(* IEC 61131-3 sources: Caravan/Archiv/12-04-19/Stations/Terminal/HMI/Network/IPCONF_IPConfigHMI, 1 file *)

(* ---- ONE_IPCONF_IPConfigHMI_Table.st ---- *)
#define OBJECTS_CONFIG

//Define part of class _IPConfigMain
//===========================================================================================================

#define MaxNoStations         50        // max. allowed No of stations

#define IPcfgWindowNrMsgBox   51000     // Window-Number of the Message Box

//===========================================================================================================
#include <.\LoaderItf.h>
//Define part of class _IPConfigStation
//===========================================================================================================

#define NiCmdIF_HmsWaitIF     20        // NewInst() command to IF object:
                                        // Time Delay for command work [100 ms] within the IF object

//===========================================================================================================

FUNCTION GLOBAL TAB ONE_IPCONF_IPConfigHMI
-1$UINT, 0$UINT,
0$UINT, 0$UINT,

13$UDINT,
TO_UDINT(3788417926), "_Global", 0$UINT, 14$UINT, 0$UINT,
TO_UDINT(1245802338), "_IPConfigIF", 1$UINT, 1$UINT, 1$UINT,
TO_UDINT(4058854491), "_IPConfigMain", 1$UINT, 2$UINT, 1$UINT,
TO_UDINT(148468755), "_IPConfigStation", 1$UINT, 2$UINT, 2$UINT,
TO_UDINT(4101473903), "_SearchUsbFiletoReset", 1$UINT, 0$UINT, 1$UINT,
TO_UDINT(2550379949), "Client_Splitter_10", 1$UINT, 2$UINT, 1$UINT,
TO_UDINT(1524808134), "Client_Splitter_Base", 1$UINT, 1$UINT, 0$UINT,
TO_UDINT(2225119864), "MerkerEx", 1$UINT, 21$UINT, 0$UINT,
TO_UDINT(3068426329), "NetworkConfig", 1$UINT, 31$UINT, 0$UINT,
TO_UDINT(933570811), "RAMex", 1$UINT, 17$UINT, 1$UINT,
TO_UDINT(2898603620), "StringInternal", 1$UINT, 82$UINT, 0$UINT,
TO_UDINT(2408581120), "StringRAM", 1$UINT, 10$UINT, 1$UINT,
TO_UDINT(3232495061), "VirtualBaseInit", 1$UINT, 3$UINT, 0$UINT,

_NO_ATTR, TO_UDINT(539668140), "_IPCONFIGIF1",

_NO_ATTR, TO_UDINT(2140441343), "_IPCONFIGMAIN1",

_NO_ATTR, TO_UDINT(2426501803), "_IPCONFIGSTATIONHMI_IF1",
_NO_ATTR, TO_UDINT(825335666), "_IPCONFIGSTATIONMC1_IF1",

_NO_ATTR, TO_UDINT(1579541752), "_SEARCHUSBFILETORESET1",

_NO_ATTR, TO_UDINT(723727191), "CLIENT_SPLITTER_101",

1$UINT, TO_UDINT(935727435), "USBSEARCHFILENAME1\DATABUFFER",

_NO_ATTR, TO_UDINT(2825064086), "USBSEARCHFILENAME1",

//Internal connections
0$UDINT,
1$UDINT,
TO_UDINT(7), "DataBuffer", TO_UDINT(6),
0$UDINT,
9$UDINT,
TO_UDINT(2), "_IPConfigMain", TO_UDINT(1), "Server0",
TO_UDINT(2), "_IPConfigIF", TO_UDINT(0), "ClassSvr",
TO_UDINT(3), "_IPConfigMain", TO_UDINT(1), "Server0",
TO_UDINT(4), "FilePathName", TO_UDINT(7), "Data",
TO_UDINT(4), "OutResetCmd", TO_UDINT(5), "To_Splitt",
TO_UDINT(5), "Ch6", TO_UDINT(3), "ExtResetCmd",
TO_UDINT(5), "Ch9", TO_UDINT(2), "ExtResetCmd",
TO_UDINT(5), "Ch10", TO_UDINT(0), "ExtResetCmd",
TO_UDINT(7), "DataBuffer", TO_UDINT(6), "m_udLength",

//Initialization values
0$UDINT,
13$UDINT,
TO_UDINT(0), "Interface", TO_UDINT(1),//|IPCONF_IPConfigHMI._IPConfigIF1.Interface;
TO_UDINT(1), "ActWindow", TO_UDINT(0),//|IPCONF_IPConfigHMI._IPConfigMain1.ActWindow;
TO_UDINT(1), "ChangeIsActive", TO_UDINT(0),//|IPCONF_IPConfigHMI._IPConfigMain1.ChangeIsActive;
TO_UDINT(2), "Timeout", TO_UDINT(30),//|IPCONF_IPConfigHMI._IPConfigStationHMI_IF1.Timeout;
TO_UDINT(2), "IsInternalIF", TO_UDINT(1),//|IPCONF_IPConfigHMI._IPConfigStationHMI_IF1.IsInternalIF;
TO_UDINT(2), "IsMMCommIF", TO_UDINT(1),//|IPCONF_IPConfigHMI._IPConfigStationHMI_IF1.IsMMCommIF;
TO_UDINT(2), "MMisOnline", TO_UDINT(0),//|IPCONF_IPConfigHMI._IPConfigStationHMI_IF1.MMisOnline;
TO_UDINT(3), "Timeout", TO_UDINT(30),//|IPCONF_IPConfigHMI._IPConfigStationMC1_IF1.Timeout;
TO_UDINT(3), "IsInternalIF", TO_UDINT(0),//|IPCONF_IPConfigHMI._IPConfigStationMC1_IF1.IsInternalIF;
TO_UDINT(3), "IsMMCommIF", TO_UDINT(1),//|IPCONF_IPConfigHMI._IPConfigStationMC1_IF1.IsMMCommIF;
TO_UDINT(3), "MMisOnline", TO_UDINT(0),//|IPCONF_IPConfigHMI._IPConfigStationMC1_IF1.MMisOnline;
TO_UDINT(6), "ThreadSafe", TO_UDINT(0),//|IPCONF_IPConfigHMI.UsbSearchFileName1\DataBuffer.ThreadSafe;
TO_UDINT(7), "SingleRealloc", TO_UDINT(1),//|IPCONF_IPConfigHMI.UsbSearchFileName1.SingleRealloc;

//Symbolic initialization values
0$UDINT,
0$UDINT,

//Initialization of string values
0$UDINT,
0$UDINT,

//Configuration of tasks (RealTime, Cyclic, Background)
0$UDINT,
0$UDINT,

0$UDINT,
0$UDINT,

0$UDINT,
4$UDINT,
TO_UDINT(0), (100)$UDINT, 4194303$DINT, 	//_IPCONFIGIF1
TO_UDINT(2), (100)$UDINT, 4194303$DINT, 	//_IPCONFIGSTATIONHMI_IF1
TO_UDINT(3), (100)$UDINT, 4194303$DINT, 	//_IPCONFIGSTATIONMC1_IF1
TO_UDINT(4), (1000)$UDINT, 4194303$DINT, 	//_SEARCHUSBFILETORESET1

//External connections
0$UDINT,
3$UDINT,
TO_UDINT(1), "Lse", C_DIR, TO_UDINT(299963966), "Lse","Lse",
TO_UDINT(1), "ActWindow", C_DIR, TO_UDINT(2925151108), "GlobalScreen1","ActWindow",
TO_UDINT(1), "ChangeIsActive", C_DIR, TO_UDINT(2516610500), "STDTCPCommunicationToMC1","DeactivateCom",

//Magic internal connections
0$UDINT,
1$UDINT,
TO_UDINT(6), "UseFile", TO_UDINT(7), "UseFile",

//Configuration of timeslots of tasks (RealTime, Cyclic)
#ifdef __LSLLDR_TIMESLOTS__
0$UDINT,
0$UDINT,

0$UDINT,
0$UDINT,

#endif //__LSLLDR_TIMESLOTS__

//MultiMaster connections
#ifdef __LSLLDR_MULTIMASTER__
0$UDINT,
1$UDINT,
TO_UDINT(3), "_IPConfigIF", C_DIR, TO_UDINT(867522694), "MachineControl._IPConfigIF1mc1.ClassSvr",
#endif //__LSLLDR_MULTIMASTER__

//Configuration for task ID (RealTime, CyclicTime)
#ifdef __LSLLDR_TASKID__
"\\\\TASKS2  "
0$UDINT,
0$UDINT,

0$UDINT,
0$UDINT,

0$UDINT,
4$UDINT,
(0)$UDINT, 	//_IPCONFIGIF1
(0)$UDINT, 	//_IPCONFIGSTATIONHMI_IF1
(0)$UDINT, 	//_IPCONFIGSTATIONMC1_IF1
(0)$UDINT, 	//_SEARCHUSBFILETORESET1

#endif //__LSLLDR_TASKID__

END_FUNCTION
